FUNCTION_BLOCK AutoCycle (* CAT Function Block Type *)
  (* Standard: 61499-2 *)
  (* Version 0.0, 11/1/2026, Schneider Electric, template *)
  PACKAGE Main;
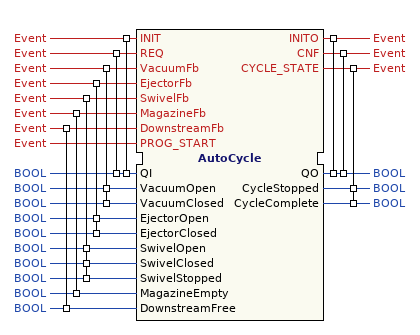
  EVENT_INPUT
    INIT WITH QI; (* Initialization Request *)
    REQ WITH QI; (* Normal Execution Request *)
    VacuumFb WITH VacuumOpen, VacuumClosed;
    EjectorFb WITH EjectorOpen, EjectorClosed;
    SwivelFb WITH SwivelOpen, SwivelClosed, SwivelStopped;
    MagazineFb WITH MagazineEmpty;
    DownstreamFb WITH DownstreamFree;
    PROG_START; (* Programmatic cycle start request *)
  END_EVENT
  EVENT_OUTPUT
    INITO WITH QO; (* Initialization Confirm *)
    CNF WITH QO; (* Execution Confirmation *)
    CYCLE_STATE WITH CycleStopped, CycleComplete; (* Sequence stopped/completed state update *)
  END_EVENT
  VAR_INPUT
    QI : BOOL; (* Input event qualifier *)
    VacuumOpen : BOOL;
    VacuumClosed : BOOL;
    EjectorOpen : BOOL;
    EjectorClosed : BOOL;
    SwivelOpen : BOOL;
    SwivelClosed : BOOL;
    SwivelStopped : BOOL;
    MagazineEmpty : BOOL;
    DownstreamFree : BOOL;
  END_VAR
  VAR_OUTPUT
    QO : BOOL; (* Output event qualifier *)
    CycleStopped : BOOL; (* TRUE when CycleSeq is Stopped *)
    CycleComplete : BOOL; (* TRUE when CycleSeq is Completed *)
  END_VAR
  FBS
    CycleSeq : SeqHead(PermStart := TRUE);
    AC1_TakeOver : SeqStep(TransStepId := 2);
    AC2_WaitDownstream : SeqStep(TransStepId := 3);
    AC3_CheckMagazine : SeqStep(TransStepId := 4);
    AC4_Eject : SeqStep(TransStepId := 5);
    AC5_EjectorBack : SeqStep(TransStepId := 6);
    AC6_ArmToMagazine : SeqStep(TransStepId := 7);
    AC7_PickUp : SeqStep(TransStepId := 8);
    AC8_Carry : SeqStep(TransStepId := 9);
    AC9_DropOff : SeqStep(TransStepId := 10);
    AC10_ParkToMag : SeqStep(TransStepId := 11);
    AC11_ParkOffMag : SeqStep(TransStepId := 12);
    AC12_ParkStop : SeqStep(TransStepId := 13);
    AC_End : SeqTerminate;
    Consts : ANY2ANY_25FC8D56FEEDC9B5(IN1 := TRUE, IN2 := 1, IN3 := 2, IN4 := 0); {SET_ATTRIBUTE(Configuration.GenericFBType.InterfaceParams, Runtime.Standard#CNT:=4;IN${CNT$}:BOOL,INT,INT,INT;OUT${CNT$}:VTQBOOL,VTQINT,VTQINT,VTQINT)}
    OwnerFb : SYMLINKMULTIVARDST_105A0442B8CC61A96(NAME1 := 'RES0.Distribution.Vacuum.sc.progLocal', NAME2 := 'RES0.Distribution.Ejector.sc.progLocal', NAME3 := 'RES0.Distribution.BlowOff.sc.progLocal', QI := TRUE); {SET_ATTRIBUTE(Configuration.GenericFBType.InterfaceParams, Runtime.System#I:=3;VALUE${I$}:VTQBOOL,VTQBOOL,VTQBOOL)}
    TakeOverCmd : SYMLINKMULTIVARSRC_32F0FE5D67925F10(QI := TRUE, NAME1 := 'RES0.Distribution.Vacuum.sc.progLocalSel', NAME2 := 'RES0.Distribution.Ejector.sc.progLocalSel', NAME3 := 'RES0.Distribution.Swivel.sc.progLocalSel', NAME4 := 'RES0.Distribution.BlowOff.sc.progLocalSel'); {SET_ATTRIBUTE(Configuration.GenericFBType.InterfaceParams, Runtime.System#I:=4;VALUE${I$}:VTQBOOL,VTQBOOL,VTQBOOL,VTQBOOL)}
    AllLocal : AND_550FE6D62F509EB3; {SET_ATTRIBUTE(Configuration.GenericFBType.InterfaceParams, Runtime.Standard#CNT:=3;OUT:BOOL)}
    MagOk : NOT_42C76073DCEB1A7A; {SET_ATTRIBUTE(Configuration.GenericFBType.InterfaceParams, Runtime.Standard#CNT:=1;OUT${CNT$}:BOOL)}
    ArmOffMag : NOT_42C76073DCEB1A7A; {SET_ATTRIBUTE(Configuration.GenericFBType.InterfaceParams, Runtime.Standard#CNT:=1;OUT${CNT$}:BOOL)}
    SwivelOutCmd : SYMLINKMULTIVARSRC_18556BCA74EA878F1(QI := TRUE, NAME1 := 'RES0.Distribution.Swivel.sc.lsp'); {SET_ATTRIBUTE(Configuration.GenericFBType.InterfaceParams, Runtime.System#I:=1;VALUE${I$}:VTQINT)}
    SwivelHomeCmd : SYMLINKMULTIVARSRC_18556BCA74EA878F1(QI := TRUE, NAME1 := 'RES0.Distribution.Swivel.sc.lsp'); {SET_ATTRIBUTE(Configuration.GenericFBType.InterfaceParams, Runtime.System#I:=1;VALUE${I$}:VTQINT)}
    BlowOnCmd : SYMLINKMULTIVARSRC_18556BCA74EA878F1(QI := TRUE, NAME1 := 'RES0.Distribution.BlowOff.sc.lsp'); {SET_ATTRIBUTE(Configuration.GenericFBType.InterfaceParams, Runtime.System#I:=1;VALUE${I$}:VTQINT)}
    EjectorBackCmd : SYMLINKMULTIVARSRC_18556BCA74EA878F1(QI := TRUE, NAME1 := 'RES0.Distribution.Ejector.sc.lsp'); {SET_ATTRIBUTE(Configuration.GenericFBType.InterfaceParams, Runtime.System#I:=1;VALUE${I$}:VTQINT)}
    VacuumOnCmd : SYMLINKMULTIVARSRC_18556BCA74EA878F1(QI := TRUE, NAME1 := 'RES0.Distribution.Vacuum.sc.lsp'); {SET_ATTRIBUTE(Configuration.GenericFBType.InterfaceParams, Runtime.System#I:=1;VALUE${I$}:VTQINT)}
    VacuumOffCmd : SYMLINKMULTIVARSRC_18556BCA74EA878F1(QI := TRUE, NAME1 := 'RES0.Distribution.Vacuum.sc.lsp'); {SET_ATTRIBUTE(Configuration.GenericFBType.InterfaceParams, Runtime.System#I:=1;VALUE${I$}:VTQINT)}
    EjectCmd : SYMLINKMULTIVARSRC_18556BCA74EA878F1(QI := TRUE, NAME1 := 'RES0.Distribution.Ejector.sc.lsp'); {SET_ATTRIBUTE(Configuration.GenericFBType.InterfaceParams, Runtime.System#I:=1;VALUE${I$}:VTQINT)}
    BlowOffCmd : SYMLINKMULTIVARSRC_18556BCA74EA878F1(QI := TRUE, NAME1 := 'RES0.Distribution.BlowOff.sc.lsp'); {SET_ATTRIBUTE(Configuration.GenericFBType.InterfaceParams, Runtime.System#I:=1;VALUE${I$}:VTQINT)}
    SwivelStopCmd : SYMLINKMULTIVARSRC_18556BCA74EA878F1(QI := TRUE, NAME1 := 'RES0.Distribution.Swivel.sc.lsp'); {SET_ATTRIBUTE(Configuration.GenericFBType.InterfaceParams, Runtime.System#I:=1;VALUE${I$}:VTQINT)}
  END_FBS
  EVENT_CONNECTIONS
    INIT TO Consts.REQ;
    Consts.CNF TO TakeOverCmd.INIT;
    Consts.CNF TO OwnerFb.INIT;
    Consts.CNF TO SwivelOutCmd.INIT;
    Consts.CNF TO SwivelHomeCmd.INIT;
    Consts.CNF TO EjectCmd.INIT;
    Consts.CNF TO EjectorBackCmd.INIT;
    Consts.CNF TO VacuumOnCmd.INIT;
    Consts.CNF TO VacuumOffCmd.INIT;
    Consts.CNF TO BlowOnCmd.INIT;
    Consts.CNF TO BlowOffCmd.INIT;
    Consts.CNF TO SwivelStopCmd.INIT;
    Consts.CNF TO CycleSeq.REQ_PERM;
    AC1_TakeOver.STEP_ENTER TO TakeOverCmd.REQ;
    TakeOverCmd.CNF TO AllLocal.REQ;
    OwnerFb.CNF TO AllLocal.REQ;
    MagazineFb TO MagOk.REQ;
    AllLocal.CNF TO AC1_TakeOver.TRANS_REQ;
    AC2_WaitDownstream.STEP_ENTER TO AC2_WaitDownstream.TRANS_REQ;
    DownstreamFb TO AC2_WaitDownstream.TRANS_REQ;
    AC3_CheckMagazine.STEP_ENTER TO MagOk.REQ;
    MagOk.CNF TO AC3_CheckMagazine.TRANS_REQ;
    AC4_Eject.STEP_ENTER TO EjectCmd.REQ;
    EjectCmd.CNF TO AC4_Eject.TRANS_REQ;
    EjectorFb TO AC4_Eject.TRANS_REQ;
    AC6_ArmToMagazine.STEP_ENTER TO SwivelHomeCmd.REQ;
    SwivelHomeCmd.CNF TO AC6_ArmToMagazine.TRANS_REQ;
    SwivelFb TO AC6_ArmToMagazine.TRANS_REQ;
    AC7_PickUp.STEP_ENTER TO VacuumOnCmd.REQ;
    VacuumOnCmd.CNF TO AC7_PickUp.TRANS_REQ;
    VacuumFb TO AC7_PickUp.TRANS_REQ;
    AC5_EjectorBack.STEP_ENTER TO EjectorBackCmd.REQ;
    EjectorBackCmd.CNF TO AC5_EjectorBack.TRANS_REQ;
    EjectorFb TO AC5_EjectorBack.TRANS_REQ;
    AC8_Carry.STEP_ENTER TO SwivelOutCmd.REQ;
    SwivelOutCmd.CNF TO AC8_Carry.TRANS_REQ;
    SwivelFb TO AC8_Carry.TRANS_REQ;
    AC9_DropOff.STEP_ENTER TO VacuumOffCmd.REQ;
    AC9_DropOff.STEP_ENTER TO BlowOnCmd.REQ;
    AC9_DropOff.STEP_LEAVE TO BlowOffCmd.REQ;
    VacuumOffCmd.CNF TO AC9_DropOff.TRANS_REQ;
    VacuumFb TO AC9_DropOff.TRANS_REQ;
    AC10_ParkToMag.STEP_ENTER TO SwivelHomeCmd.REQ;
    SwivelHomeCmd.CNF TO AC10_ParkToMag.TRANS_REQ;
    SwivelFb TO AC10_ParkToMag.TRANS_REQ;
    AC11_ParkOffMag.STEP_ENTER TO SwivelOutCmd.REQ;
    SwivelOutCmd.CNF TO ArmOffMag.REQ;
    SwivelFb TO ArmOffMag.REQ;
    ArmOffMag.CNF TO AC11_ParkOffMag.TRANS_REQ;
    AC12_ParkStop.STEP_ENTER TO SwivelStopCmd.REQ;
    SwivelStopCmd.CNF TO AC12_ParkStop.TRANS_REQ;
    SwivelFb TO AC12_ParkStop.TRANS_REQ;
    PROG_START TO CycleSeq.START;
    CycleSeq.STATE_IND TO CYCLE_STATE;
  END_CONNECTIONS
  DATA_CONNECTIONS
    Consts.OUT1 TO TakeOverCmd.VALUE1;
    Consts.OUT1 TO TakeOverCmd.VALUE2;
    Consts.OUT1 TO TakeOverCmd.VALUE3;
    Consts.OUT1 TO TakeOverCmd.VALUE4;
    Consts.OUT2 TO SwivelOutCmd.VALUE1;
    Consts.OUT2 TO EjectCmd.VALUE1;
    Consts.OUT2 TO VacuumOnCmd.VALUE1;
    Consts.OUT2 TO BlowOnCmd.VALUE1;
    Consts.OUT3 TO SwivelHomeCmd.VALUE1;
    Consts.OUT3 TO EjectorBackCmd.VALUE1;
    Consts.OUT3 TO VacuumOffCmd.VALUE1;
    Consts.OUT4 TO BlowOffCmd.VALUE1;
    Consts.OUT4 TO SwivelStopCmd.VALUE1;
    OwnerFb.VALUE1 TO AllLocal.IN1;
    OwnerFb.VALUE2 TO AllLocal.IN2;
    OwnerFb.VALUE3 TO AllLocal.IN3;
    MagazineEmpty TO MagOk.IN1;
    AllLocal.OUT TO AC1_TakeOver.Exceeded;
    DownstreamFree TO AC2_WaitDownstream.Exceeded;
    MagOk.OUT1 TO AC3_CheckMagazine.Exceeded;
    EjectorOpen TO AC4_Eject.Exceeded;
    SwivelClosed TO AC6_ArmToMagazine.Exceeded;
    VacuumOpen TO AC7_PickUp.Exceeded;
    EjectorClosed TO AC5_EjectorBack.Exceeded;
    SwivelOpen TO AC8_Carry.Exceeded;
    VacuumClosed TO AC9_DropOff.Exceeded;
    SwivelClosed TO AC10_ParkToMag.Exceeded;
    SwivelClosed TO ArmOffMag.IN1;
    ArmOffMag.OUT1 TO AC11_ParkOffMag.Exceeded;
    SwivelStopped TO AC12_ParkStop.Exceeded;
    CycleSeq.SeqStopped TO CycleStopped;
    CycleSeq.SeqComplete TO CycleComplete;
  END_CONNECTIONS
  ADAPTER_CONNECTIONS
    CycleSeq.ISeqChain TO AC1_TakeOver.ISeqChainIn;
    AC1_TakeOver.ISeqChainOut TO AC2_WaitDownstream.ISeqChainIn;
    AC2_WaitDownstream.ISeqChainOut TO AC3_CheckMagazine.ISeqChainIn;
    AC3_CheckMagazine.ISeqChainOut TO AC4_Eject.ISeqChainIn;
    AC4_Eject.ISeqChainOut TO AC5_EjectorBack.ISeqChainIn;
    AC5_EjectorBack.ISeqChainOut TO AC6_ArmToMagazine.ISeqChainIn;
    AC6_ArmToMagazine.ISeqChainOut TO AC7_PickUp.ISeqChainIn;
    AC7_PickUp.ISeqChainOut TO AC8_Carry.ISeqChainIn;
    AC8_Carry.ISeqChainOut TO AC9_DropOff.ISeqChainIn;
    AC9_DropOff.ISeqChainOut TO AC10_ParkToMag.ISeqChainIn;
    AC10_ParkToMag.ISeqChainOut TO AC11_ParkOffMag.ISeqChainIn;
    AC11_ParkOffMag.ISeqChainOut TO AC12_ParkStop.ISeqChainIn;
    AC12_ParkStop.ISeqChainOut TO AC_End.ISeqChainIn;
  END_CONNECTIONS
END_FUNCTION_BLOCK
